(* IEC 61131-3 sources: 2026_Projet_YGO_ExcavatriceDragage/ARCHIVES/Code/PLC_TESTS, 2 files *)

(* ---- GVL_PLC_Tests_Const.st ---- *)
(* ═══════════════════════════════════════════════════════════════
   🧪 GVL_PLC_Tests_Const — Constantes de dimensionnement
   ───────────────────────────────────────────────────────────────
   🎯 Rôle : Définit les tailles limites des tables de tests
      pour l'orchestrateur et le moteur de tests.
   ═══════════════════════════════════════════════════════════════ *)

{attribute 'qualified_only'}
VAR_GLOBAL CONSTANT
    MaxTestCases     : INT := 8;    // par suite
    MaxSteps         : INT := 128;  // par suite, table PLATE ; WINCH-CORE-01 ajoute les étapes 65..111
    MaxChecks        : INT := 64;   // CheckTable par suite
    MaxChecksPerStep : INT := 10;
    MaxInvariants    : INT := 4;    // actifs en parallèle
    MaxProbeBool     : INT := 32;
    MaxProbeDint     : INT := 16;    // INT/WORD/étapes séquenceur → conversion au câblage (WORD_TO_DINT)
    MaxProbeReal     : INT := 16;    // analogiques + TIME → REAL ms
    MaxAnalogStims   : INT := 4;    // instances FB_TestStimulus par suite
    MaxSeqValues     : INT := 8;    // plus gros poste mémoire par stim
    TaskCycleMs      : INT := 10;   // MainTask — base des mesures en cycles
    MaxSuiteDurationMs : DINT := 180000; // 🛡️ garde-fou orchestrateur : 3 min maximum par suite
    MaxTestEvents    : INT := 32;   // journal circulaire des événements
    SuiteSafety      : INT := 1;    // index de suite (Cmd.RunSuite)
    SuiteTranslation : INT := 2;    // index de suite Translation M3 (Cmd.RunSuite)
    SuiteBucket      : INT := 3;    // index de suite Bucket (Cmd.RunSuite)
    SuiteEncoder     : INT := 4;    // index de suite Codeurs/Homing nominal (Cmd.RunSuite)
    SuiteModes       : INT := 5;    // index de suite Modes/Homme-mort, post-suppression IHM_MANU (Cmd.RunSuite)
    SuiteHeartbeat   : INT := 6;    // index de suite Heartbeat IHM↔PLC (Cmd.RunSuite)
    SuiteSupervision : INT := 8;    // index Supervision/Persistance config — 7 = Framework Validation
END_VAR

(* ---- FB_TestSequencer.st ---- *)
FUNCTION_BLOCK FB_TestSequencer
VAR_INPUT
    Start       : BOOL;              // Front : lance la suite
    Abort       : BOOL;              // Niveau : arrêt immédiat propre
    CaseId      : INT;               // 0=tous ; 1..MaxTestCases=cas ciblé
END_VAR
VAR_IN_OUT                           // 🔗 zéro copie
    StepTable      : ARRAY[1..GVL_PLC_Tests_Const.MaxSteps]      OF ST_TestStepConfig;
    CheckTable     : ARRAY[1..GVL_PLC_Tests_Const.MaxChecks]     OF ST_TestCheckConfig;
    CaseTable      : ARRAY[1..GVL_PLC_Tests_Const.MaxTestCases]  OF ST_TestCaseConfig;
    InvariantTable : ARRAY[1..GVL_PLC_Tests_Const.MaxInvariants] OF ST_TestInvariantConfig;
    ProbeBool      : ARRAY[1..GVL_PLC_Tests_Const.MaxProbeBool]  OF BOOL;
    ProbeDint      : ARRAY[1..GVL_PLC_Tests_Const.MaxProbeDint]  OF DINT;
    ProbeReal      : ARRAY[1..GVL_PLC_Tests_Const.MaxProbeReal]  OF REAL;
    Report         : ST_TestSuiteReport;
END_VAR
VAR_OUTPUT
    Busy                : BOOL;
    Done                : BOOL;
    AnyFailed           : BOOL;
    ConfigError         : BOOL;      // 🔒 Table invalide -> refus de lancer
    ConfigErrorStepId   : INT;
    ConfigErrorCheckIdx : INT;
    TerminalState       : E_TestTerminalState;
    ErrorCode           : INT;
    ErrorMessage        : STRING(160);
    CurrentStepId       : INT;
    ActiveStimulusId    : INT;       // ⚡ consommé par le domaine
    StepElapsed         : TIME;      // Pour l'IHM
END_VAR
VAR
    StartTrig           : R_TRIG;
    StepTimer           : TON;
    DwellTimer          : TON;
    Checks              : ARRAY[1..GVL_PLC_Tests_Const.MaxChecksPerStep] OF FB_TestCheck;
    InvChecks           : ARRAY[1..GVL_PLC_Tests_Const.MaxInvariants]    OF FB_TestCheck;
    InvArmed            : ARRAY[1..GVL_PLC_Tests_Const.MaxInvariants]    OF BOOL;

    // Variables de contrôle internes
    StepStarted         : BOOL;
    CurrentCaseId       : INT;
    Idx                 : INT;
    Jdx                 : INT;
    Kdx                 : INT;
    Valid               : BOOL;

    // 🔧 REX : locaux remontés depuis des blocs VAR imbriqués dans le corps
    AllChecksPassed     : BOOL;
    AnyCheckFailed      : BOOL;
    FailedCheckIdxLocal : INT;
    FailReasonLocal     : E_TestFailReason;
    ObsBoolLocal        : BOOL;
    ObsDintLocal        : DINT;
    ObsRealLocal        : REAL;
    NeverDuringPassed   : BOOL;
    SuiteAllPassed      : BOOL;
    FirstFailedCase     : INT;
    CaseIdx             : INT;
    CaseStartStep       : INT;
    CaseStep            : INT;
    CaseWalkCount       : INT;
    CaseOk              : BOOL;
    CaseExecuted        : BOOL;
    CaseFailedStep      : INT;
    CaseDuration        : TIME;
    CaseFailReason      : E_TestFailReason;

    // 🏷️ Construction de Report.FailureSummary (1 ligne lisible, tous les cas en échec)
    ReasonText          : STRING(20);
    EntryText           : STRING(80);
    FirstStepLocal      : INT;
    RequestedCaseId     : INT;
END_VAR
// === IMPLEMENTATION ===
StartTrig(CLK := Start);

// 1. Validation de la configuration sur front de Start
IF StartTrig.Q THEN
    ConfigError := FALSE;
    ConfigErrorStepId := 0;
    ConfigErrorCheckIdx := 0;
    TerminalState := E_TestTerminalState.TEST_TERMINAL_NONE;
    ErrorCode := 0;
    ErrorMessage := '';

    // 🛡️ Résolution interne CaseId → première étape, jamais d'étape exposée.
    RequestedCaseId := CaseId;
    IF CaseId < 0 OR CaseId > GVL_PLC_Tests_Const.MaxTestCases THEN
        ConfigError := TRUE;
        ConfigErrorStepId := CaseId;
        ErrorCode := 1001;
        ErrorMessage := 'CaseId hors limites';
        FirstStepLocal := 0;
    ELSIF CaseId = 0 THEN
        FirstStepLocal := CaseTable[1].FirstStep;
    ELSE
        FirstStepLocal := CaseTable[CaseId].FirstStep;
    END_IF;
    IF NOT ConfigError THEN
        IF FirstStepLocal < 1 OR FirstStepLocal > GVL_PLC_Tests_Const.MaxSteps THEN
            ConfigError := TRUE;
            ConfigErrorStepId := FirstStepLocal;
            ErrorCode := 1001;
            ErrorMessage := 'CaseTable.FirstStep hors limites';
        END_IF;
    END_IF;

    // Validation des étapes
    FOR Idx := 1 TO GVL_PLC_Tests_Const.MaxSteps DO
        IF StepTable[Idx].CaseId > 0 THEN
            // Vérification des NextOn
            IF StepTable[Idx].NextOnPass < 0 OR StepTable[Idx].NextOnPass > GVL_PLC_Tests_Const.MaxSteps THEN
                ConfigError := TRUE;
                ConfigErrorStepId := Idx;
            ELSIF StepTable[Idx].NextOnFail < 0 OR StepTable[Idx].NextOnFail > GVL_PLC_Tests_Const.MaxSteps THEN
                ConfigError := TRUE;
                ConfigErrorStepId := Idx;
            END_IF;

            // Vérification du Timeout
            IF StepTable[Idx].TimeoutPT <= T#0s THEN
                // Sauf si tous les checks de cette étape sont NEVER_DURING, mais restons stricts : TimeoutPT requis
                ConfigError := TRUE;
                ConfigErrorStepId := Idx;
            END_IF;

            // Vérification des Checks indexés par l'étape
            FOR Jdx := 1 TO GVL_PLC_Tests_Const.MaxChecksPerStep DO
                Kdx := StepTable[Idx].CheckIdx[Jdx];
                IF Kdx > 0 THEN
                    IF Kdx > GVL_PLC_Tests_Const.MaxChecks THEN
                        ConfigError := TRUE;
                        ConfigErrorStepId := Idx;
                        ConfigErrorCheckIdx := Kdx;
                    ELSE
                        // Validation de la sonde associée au check
                        CASE CheckTable[Kdx].Kind OF
                            E_TestCheckKind.BOOL_EQUAL, E_TestCheckKind.BOOL_RISING, E_TestCheckKind.BOOL_FALLING:
                                IF CheckTable[Kdx].ProbeIdx < 1 OR CheckTable[Kdx].ProbeIdx > GVL_PLC_Tests_Const.MaxProbeBool THEN
                                    ConfigError := TRUE;
                                    ConfigErrorStepId := Idx;
                                    ConfigErrorCheckIdx := Kdx;
                                END_IF;
                            E_TestCheckKind.DINT_EQUAL, E_TestCheckKind.DINT_NOT_EQUAL, E_TestCheckKind.DINT_IN_RANGE,
                            E_TestCheckKind.WORD_MASK_ALL, E_TestCheckKind.WORD_MASK_ANY, E_TestCheckKind.WORD_MASK_NONE:
                                IF CheckTable[Kdx].ProbeIdx < 1 OR CheckTable[Kdx].ProbeIdx > GVL_PLC_Tests_Const.MaxProbeDint THEN
                                    ConfigError := TRUE;
                                    ConfigErrorStepId := Idx;
                                    ConfigErrorCheckIdx := Kdx;
                                END_IF;
                            E_TestCheckKind.REAL_IN_RANGE:
                                IF CheckTable[Kdx].ProbeIdx < 1 OR CheckTable[Kdx].ProbeIdx > GVL_PLC_Tests_Const.MaxProbeReal THEN
                                    ConfigError := TRUE;
                                    ConfigErrorStepId := Idx;
                                    ConfigErrorCheckIdx := Kdx;
                                END_IF;
                        END_CASE;
                    END_IF;
                END_IF;
            END_FOR;
        END_IF;
    END_FOR;

    // 🛡️ ConfigError doit toujours produire Done + un état terminal.
    IF ConfigError THEN
        Busy := FALSE;
        Done := TRUE;
        AnyFailed := TRUE;
        ActiveStimulusId := 0;
        CurrentStepId := 0;
        StepElapsed := T#0s;
        TerminalState := E_TestTerminalState.TEST_TERMINAL_CONFIG_ERROR;
        Report.InProgress := FALSE;
        Report.RunCounter := Report.RunCounter + 1;
        Report.AllPassed := FALSE;
        Report.AnyFailed := TRUE;
        Report.Aborted := FALSE;
        Report.TerminalState := TerminalState;
        IF ErrorCode = 0 THEN
            ErrorCode := 1002;
            ErrorMessage := 'Table de test invalide';
        END_IF;
        Report.ErrorCode := ErrorCode;
        Report.ErrorMessage := ErrorMessage;
        Report.FailureSummary := CONCAT('CONFIG_ERROR step ', INT_TO_STRING(ConfigErrorStepId));
        RETURN;
    END_IF;
END_IF;

// 2. Abort (Niveau, priorité absolue)
IF Abort THEN
    IF Busy THEN
        Report.InProgress := FALSE;
        Report.Aborted := TRUE;
        Report.AnyFailed := TRUE;

        // Enregistrement de l'échec de l'étape courante
        IF CurrentStepId >= 1 AND CurrentStepId <= GVL_PLC_Tests_Const.MaxSteps THEN
            Report.Steps[CurrentStepId].Executed := TRUE;
            Report.Steps[CurrentStepId].Passed := FALSE;
            Report.Steps[CurrentStepId].FailReason := E_TestFailReason.FAIL_ABORTED;
            Report.Steps[CurrentStepId].Duration := StepElapsed;
        END_IF;

        // Échec du cas de test en cours
        IF CurrentCaseId >= 1 AND CurrentCaseId <= GVL_PLC_Tests_Const.MaxTestCases THEN
            Report.Cases[CurrentCaseId].Ok := FALSE;
            Report.Cases[CurrentCaseId].FailReason := E_TestFailReason.FAIL_ABORTED;
        END_IF;

        Busy := FALSE;
        Done := TRUE;
        AnyFailed := TRUE;
        TerminalState := E_TestTerminalState.TEST_TERMINAL_ABORTED;
        Report.TerminalState := TerminalState;
    END_IF;
    ActiveStimulusId := 0;
    StepStarted := FALSE;
    RETURN;
END_IF;

// 3. Démarrage de la suite
IF StartTrig.Q AND NOT ConfigError THEN
    Busy := TRUE;
    Done := FALSE;
    AnyFailed := FALSE;
    CurrentStepId := FirstStepLocal;
    StepStarted := FALSE;

    // RAZ Rapport
    Report.InProgress := TRUE;
    Report.AllPassed := FALSE;
    Report.AnyFailed := FALSE;
    Report.Aborted := FALSE;
    Report.TerminalState := E_TestTerminalState.TEST_TERMINAL_NONE;
    Report.ErrorCode := 0;
    Report.ErrorMessage := '';
    Report.FailedTestCase := 0;
    Report.CurrentStepId := FirstStepLocal;
    IF CurrentStepId >= 1 AND CurrentStepId <= GVL_PLC_Tests_Const.MaxSteps THEN
        Report.CurrentCaseId := StepTable[CurrentStepId].CaseId;
    ELSE
        Report.CurrentCaseId := 0;
    END_IF;
    Report.Duration := T#0s;
    Report.RunCounter := Report.RunCounter + 1;

    FOR Idx := 1 TO GVL_PLC_Tests_Const.MaxSteps DO
        Report.Steps[Idx].Executed := FALSE;
        Report.Steps[Idx].Passed := FALSE;
        Report.Steps[Idx].FailReason := E_TestFailReason.FAIL_NONE;
        Report.Steps[Idx].FailedCheckIdx := 0;
        Report.Steps[Idx].FailedInvariantId := 0;
        Report.Steps[Idx].Duration := T#0s;
    END_FOR;

    FOR Idx := 1 TO GVL_PLC_Tests_Const.MaxTestCases DO
        Report.Cases[Idx].Executed := FALSE;
        Report.Cases[Idx].Ok := FALSE;
        Report.Cases[Idx].FailedStepId := 0;
        Report.Cases[Idx].FailReason := E_TestFailReason.FAIL_NONE;
        Report.Cases[Idx].Duration := T#0s;
    END_FOR;

    // RAZ Invariants
    FOR Idx := 1 TO GVL_PLC_Tests_Const.MaxInvariants DO
        InvArmed[Idx] := FALSE;
    END_FOR;
END_IF;

// 4. Moteur d'exécution principal
IF Busy THEN
    // Incrément de la durée globale du run
    Report.Duration := Report.Duration + UDINT_TO_TIME(INT_TO_UDINT(GVL_PLC_Tests_Const.TaskCycleMs));

    // Vérification des bornes de l'étape courante (0 est valide et désigne la fin)
    IF CurrentStepId <> 0 AND (CurrentStepId < 1 OR CurrentStepId > GVL_PLC_Tests_Const.MaxSteps) THEN
        Busy := FALSE;
        Done := TRUE;
        AnyFailed := TRUE;
        ActiveStimulusId := 0;
        ConfigError := TRUE;
        ConfigErrorStepId := CurrentStepId;
        ErrorCode := 1003;
        ErrorMessage := 'Etape courante hors limites';
        TerminalState := E_TestTerminalState.TEST_TERMINAL_CONFIG_ERROR;
        Report.InProgress := FALSE;
        Report.AnyFailed := TRUE;
        Report.TerminalState := TerminalState;
        Report.ErrorCode := ErrorCode;
        Report.ErrorMessage := ErrorMessage;
        Report.FailureSummary := ErrorMessage;
        RETURN;
    END_IF;

    // 🔒 Fin automatique dès qu'un run ciblé tenterait d'entrer dans le cas suivant.
    IF CurrentStepId > 0 AND RequestedCaseId > 0 THEN
        IF StepTable[CurrentStepId].CaseId <> RequestedCaseId THEN
            CurrentStepId := 0;
            ActiveStimulusId := 0;
            StepStarted := FALSE;
        END_IF;
    END_IF;

    IF CurrentStepId > 0 THEN
    CurrentCaseId := StepTable[CurrentStepId].CaseId;
    ActiveStimulusId := StepTable[CurrentStepId].StimulusId;
    Report.CurrentStepId := CurrentStepId;
    Report.CurrentCaseId := CurrentCaseId;

    IF NOT StepStarted THEN
        StepStarted := TRUE;
        StepElapsed := T#0s;
        DwellTimer(IN := FALSE);
        StepTimer(IN := FALSE);

        // Gestion de l'armement/désarmement des invariants
        FOR Idx := 1 TO GVL_PLC_Tests_Const.MaxInvariants DO
            IF InvariantTable[Idx].ArmAtStepId = CurrentStepId THEN
                InvArmed[Idx] := TRUE;
            END_IF;
            IF InvariantTable[Idx].DisarmAtStepId = CurrentStepId THEN
                InvArmed[Idx] := FALSE;
            END_IF;
        END_FOR;
    END_IF;

    // Incrément de la durée de l'étape courante
    StepElapsed := StepElapsed + UDINT_TO_TIME(INT_TO_UDINT(GVL_PLC_Tests_Const.TaskCycleMs));

    // 4.1 Évaluation des invariants actifs
    FOR Idx := 1 TO GVL_PLC_Tests_Const.MaxInvariants DO
        IF InvArmed[Idx] THEN
            InvChecks[Idx](Config := InvariantTable[Idx].Check, Evaluate := TRUE, ProbeBool := ProbeBool, ProbeDint := ProbeDint, ProbeReal := ProbeReal);
            IF InvChecks[Idx].Failed THEN
                // Violation d'invariant -> Transition en échec immédiat
                Report.Steps[CurrentStepId].Executed := TRUE;
                Report.Steps[CurrentStepId].Passed := FALSE;
                Report.Steps[CurrentStepId].FailReason := E_TestFailReason.FAIL_INVARIANT;
                Report.Steps[CurrentStepId].FailedInvariantId := Idx;
                Report.Steps[CurrentStepId].Duration := StepElapsed;
                Report.Steps[CurrentStepId].ObservedBool := InvChecks[Idx].ObservedBool;
                Report.Steps[CurrentStepId].ObservedDint := InvChecks[Idx].ObservedDint;
                Report.Steps[CurrentStepId].ObservedReal := InvChecks[Idx].ObservedReal;

                // Désactivation de l'évaluation
                InvChecks[Idx](Config := InvariantTable[Idx].Check, Evaluate := FALSE, ProbeBool := ProbeBool, ProbeDint := ProbeDint, ProbeReal := ProbeReal);

                // Transition
                IF StepTable[CurrentStepId].FailAction = E_TestFailAction.FAIL_ABORT_SUITE THEN
                    Busy := FALSE;
                    Done := TRUE;
                    AnyFailed := TRUE;
                    ActiveStimulusId := 0;
                ELSE
                    CurrentStepId := StepTable[CurrentStepId].NextOnFail;
                    StepStarted := FALSE;
                END_IF;
                RETURN;
            END_IF;
        END_IF;
    END_FOR;

    // 4.2 Gestion de la temporisation de Dwell
    DwellTimer(IN := TRUE, PT := StepTable[CurrentStepId].DwellPT);
    IF NOT DwellTimer.Q THEN
        // En attente du Dwell, pas d'évaluation des checks d'étape
        FOR Jdx := 1 TO GVL_PLC_Tests_Const.MaxChecksPerStep DO
            Checks[Jdx](Evaluate := FALSE, ProbeBool := ProbeBool, ProbeDint := ProbeDint, ProbeReal := ProbeReal);
        END_FOR;
        RETURN;
    END_IF;

    // 4.3 Évaluation des checks d'étape
    AllChecksPassed     := TRUE;
    AnyCheckFailed      := FALSE;
    FailedCheckIdxLocal := 0;
    FailReasonLocal     := E_TestFailReason.FAIL_NONE;
    ObsBoolLocal        := FALSE;
    ObsDintLocal        := 0;
    ObsRealLocal        := 0.0;

    FOR Jdx := 1 TO GVL_PLC_Tests_Const.MaxChecksPerStep DO
        Kdx := StepTable[CurrentStepId].CheckIdx[Jdx];
        IF Kdx < 0 OR Kdx > GVL_PLC_Tests_Const.MaxChecks THEN
            ConfigError := TRUE;
            ConfigErrorStepId := CurrentStepId;
            ConfigErrorCheckIdx := Kdx;
            ErrorCode := 1006;
            ErrorMessage := 'CheckIdx runtime hors limites';
            Busy := FALSE;
            Done := TRUE;
            AnyFailed := TRUE;
            ActiveStimulusId := 0;
            TerminalState := E_TestTerminalState.TEST_TERMINAL_CONFIG_ERROR;
            RETURN;
        END_IF;
        IF Kdx > 0 THEN
            Checks[Jdx](Config := CheckTable[Kdx], Evaluate := TRUE, ProbeBool := ProbeBool, ProbeDint := ProbeDint, ProbeReal := ProbeReal);

            IF Checks[Jdx].Failed THEN
                AnyCheckFailed := TRUE;
                FailedCheckIdxLocal := Kdx;
                FailReasonLocal := Checks[Jdx].FailReason;
                ObsBoolLocal := Checks[Jdx].ObservedBool;
                ObsDintLocal := Checks[Jdx].ObservedDint;
                ObsRealLocal := Checks[Jdx].ObservedReal;
            ELSIF Checks[Jdx].Pending THEN
                AllChecksPassed := FALSE;
            END_IF;
        END_IF;
    END_FOR;

    // 4.4 Prise de verdict
    IF AnyCheckFailed THEN
        // Échec sur un check d'étape
        Report.Steps[CurrentStepId].Executed := TRUE;
        Report.Steps[CurrentStepId].Passed := FALSE;
        Report.Steps[CurrentStepId].FailReason := FailReasonLocal;
        Report.Steps[CurrentStepId].FailedCheckIdx := FailedCheckIdxLocal;
        Report.Steps[CurrentStepId].Duration := StepElapsed;
        Report.Steps[CurrentStepId].ObservedBool := ObsBoolLocal;
        Report.Steps[CurrentStepId].ObservedDint := ObsDintLocal;
        Report.Steps[CurrentStepId].ObservedReal := ObsRealLocal;

        // Reset checks
        FOR Jdx := 1 TO GVL_PLC_Tests_Const.MaxChecksPerStep DO
            Checks[Jdx](Evaluate := FALSE, ProbeBool := ProbeBool, ProbeDint := ProbeDint, ProbeReal := ProbeReal);
        END_FOR;

        IF StepTable[CurrentStepId].FailAction = E_TestFailAction.FAIL_ABORT_SUITE THEN
            Busy := FALSE;
            Done := TRUE;
            AnyFailed := TRUE;
            ActiveStimulusId := 0;
        ELSE
            CurrentStepId := StepTable[CurrentStepId].NextOnFail;
            StepStarted := FALSE;
        END_IF;
        RETURN;
    END_IF;

    StepTimer(IN := TRUE, PT := StepTable[CurrentStepId].TimeoutPT);

    IF AllChecksPassed THEN
        // Succès précoce (vérification MinPT)
        IF StepElapsed < StepTable[CurrentStepId].MinPT THEN
            // Réaction trop rapide = Échec
            Report.Steps[CurrentStepId].Executed := TRUE;
            Report.Steps[CurrentStepId].Passed := FALSE;
            Report.Steps[CurrentStepId].FailReason := E_TestFailReason.FAIL_WINDOW_EARLY;
            Report.Steps[CurrentStepId].Duration := StepElapsed;

            // Reset checks
            FOR Jdx := 1 TO GVL_PLC_Tests_Const.MaxChecksPerStep DO
                Checks[Jdx](Evaluate := FALSE, ProbeBool := ProbeBool, ProbeDint := ProbeDint, ProbeReal := ProbeReal);
            END_FOR;

            IF StepTable[CurrentStepId].FailAction = E_TestFailAction.FAIL_ABORT_SUITE THEN
                Busy := FALSE;
                Done := TRUE;
                AnyFailed := TRUE;
                ActiveStimulusId := 0;
            ELSE
                CurrentStepId := StepTable[CurrentStepId].NextOnFail;
                StepStarted := FALSE;
            END_IF;
        ELSE
            // Validation étape OK
            Report.Steps[CurrentStepId].Executed := TRUE;
            Report.Steps[CurrentStepId].Passed := TRUE;
            Report.Steps[CurrentStepId].Duration := StepElapsed;

            // Prendre snapshot du premier check s'il existe
            IF StepTable[CurrentStepId].CheckIdx[1] > 0 THEN
                Report.Steps[CurrentStepId].ObservedBool := Checks[1].ObservedBool;
                Report.Steps[CurrentStepId].ObservedDint := Checks[1].ObservedDint;
                Report.Steps[CurrentStepId].ObservedReal := Checks[1].ObservedReal;
            END_IF;

            // Reset checks
            FOR Jdx := 1 TO GVL_PLC_Tests_Const.MaxChecksPerStep DO
                Checks[Jdx](Evaluate := FALSE, ProbeBool := ProbeBool, ProbeDint := ProbeDint, ProbeReal := ProbeReal);
            END_FOR;

            CurrentStepId := StepTable[CurrentStepId].NextOnPass;
            StepStarted := FALSE;
        END_IF;
        RETURN;
    END_IF;

    // Gestion du timeout d'étape
    IF StepTimer.Q THEN
        // Si timeout expiré, vérifions si des checks NEVER_DURING sont en attente
        NeverDuringPassed := TRUE;
        FOR Jdx := 1 TO GVL_PLC_Tests_Const.MaxChecksPerStep DO
            Kdx := StepTable[CurrentStepId].CheckIdx[Jdx];
            IF Kdx < 0 OR Kdx > GVL_PLC_Tests_Const.MaxChecks THEN
                ConfigError := TRUE;
                ConfigErrorStepId := CurrentStepId;
                ConfigErrorCheckIdx := Kdx;
                ErrorCode := 1006;
                ErrorMessage := 'CheckIdx timeout hors limites';
                Busy := FALSE;
                Done := TRUE;
                AnyFailed := TRUE;
                ActiveStimulusId := 0;
                TerminalState := E_TestTerminalState.TEST_TERMINAL_CONFIG_ERROR;
                RETURN;
            END_IF;
            IF Kdx > 0 THEN
                IF CheckTable[Kdx].Mode = E_TestCheckMode.CHECK_NEVER_DURING THEN
                    // Jamais violé pendant toute la fenêtre
                    Checks[Jdx](Evaluate := FALSE, ProbeBool := ProbeBool, ProbeDint := ProbeDint, ProbeReal := ProbeReal);
                ELSE
                    // Les autres modes auraient dû passer avant le timeout
                    NeverDuringPassed := FALSE;
                END_IF;
            END_IF;
        END_FOR;

        IF NeverDuringPassed THEN
            // Succès par non-violation
            Report.Steps[CurrentStepId].Executed := TRUE;
            Report.Steps[CurrentStepId].Passed := TRUE;
            Report.Steps[CurrentStepId].Duration := StepElapsed;

            CurrentStepId := StepTable[CurrentStepId].NextOnPass;
            StepStarted := FALSE;
        ELSE
            // Timeout classique de l'étape
            Report.Steps[CurrentStepId].Executed := TRUE;
            Report.Steps[CurrentStepId].Passed := FALSE;
            Report.Steps[CurrentStepId].FailReason := E_TestFailReason.FAIL_TIMEOUT;
            Report.Steps[CurrentStepId].Duration := StepElapsed;

            IF StepTable[CurrentStepId].FailAction = E_TestFailAction.FAIL_ABORT_SUITE THEN
                Busy := FALSE;
                Done := TRUE;
                AnyFailed := TRUE;
                ActiveStimulusId := 0;
            ELSE
                CurrentStepId := StepTable[CurrentStepId].NextOnFail;
                StepStarted := FALSE;
            END_IF;
        END_IF;

        // Reset checks
        FOR Jdx := 1 TO GVL_PLC_Tests_Const.MaxChecksPerStep DO
            Checks[Jdx](Evaluate := FALSE, ProbeBool := ProbeBool, ProbeDint := ProbeDint, ProbeReal := ProbeReal);
        END_FOR;
    END_IF;
    END_IF;
END_IF;

// 5. Agrégation des résultats en fin de suite (CurrentStepId = 0)
IF Busy AND CurrentStepId = 0 THEN
    Busy := FALSE;
    Done := TRUE;
    ActiveStimulusId := 0;
    Report.InProgress := FALSE;

    // Agrégation des cas de test
    SuiteAllPassed  := TRUE;
    FirstFailedCase := 0;

    FOR CaseIdx := 1 TO GVL_PLC_Tests_Const.MaxTestCases DO
        CaseStartStep := CaseTable[CaseIdx].FirstStep;
        IF CaseStartStep > 0 THEN
            CaseOk := TRUE;
            CaseExecuted := FALSE;
            CaseFailedStep := 0;
            CaseDuration := T#0s;
            CaseFailReason := E_TestFailReason.FAIL_NONE;

            // 🔒 Parcours borné et index validé AVANT déréférencement.
            // CODESYS peut évaluer StepTable[CaseStep] même si CaseStep=0
            // dans une condition composée : ancienne version = Access Violation CPU.
            CaseStep := CaseStartStep;
            FOR CaseWalkCount := 1 TO GVL_PLC_Tests_Const.MaxSteps DO
                IF CaseStep = 0 THEN
                    EXIT;
                END_IF;
                IF CaseStep < 1 OR CaseStep > GVL_PLC_Tests_Const.MaxSteps THEN
                    ConfigError := TRUE;
                    ConfigErrorStepId := CaseStep;
                    ErrorCode := 1004;
                    ErrorMessage := 'Agregation : etape hors limites';
                    CaseOk := FALSE;
                    EXIT;
                END_IF;
                IF StepTable[CaseStep].CaseId <> CaseIdx THEN
                    EXIT;
                END_IF;

                IF Report.Steps[CaseStep].Executed THEN
                    CaseExecuted := TRUE;
                    CaseDuration := CaseDuration + Report.Steps[CaseStep].Duration;
                    IF NOT Report.Steps[CaseStep].Passed THEN
                        CaseOk := FALSE;
                        CaseFailedStep := CaseStep;
                        CaseFailReason := Report.Steps[CaseStep].FailReason;
                        CaseStep := StepTable[CaseStep].NextOnFail;
                    ELSE
                        CaseStep := StepTable[CaseStep].NextOnPass;
                    END_IF;
                ELSE
                    CaseStep := StepTable[CaseStep].NextOnPass;
                END_IF;
            END_FOR;
            IF CaseStep <> 0 AND CaseWalkCount > GVL_PLC_Tests_Const.MaxSteps THEN
                ConfigError := TRUE;
                ConfigErrorStepId := CaseStep;
                ErrorCode := 1005;
                ErrorMessage := 'Agregation : cycle de transitions';
                CaseOk := FALSE;
            END_IF;

            Report.Cases[CaseIdx].Name := CaseTable[CaseIdx].Name; // 🏷️ Lisible directement en Watch, sans chercher l'index
            Report.Cases[CaseIdx].Executed := CaseExecuted;
            Report.Cases[CaseIdx].Ok := CaseExecuted AND CaseOk;
            Report.Cases[CaseIdx].FailedStepId := CaseFailedStep;
            Report.Cases[CaseIdx].FailReason := CaseFailReason;
            Report.Cases[CaseIdx].Duration := CaseDuration;

            IF CaseExecuted AND NOT CaseOk THEN
                SuiteAllPassed := FALSE;
                IF FirstFailedCase = 0 THEN
                    FirstFailedCase := CaseIdx;
                END_IF;
            END_IF;
        END_IF;
    END_FOR;

    Report.AllPassed := SuiteAllPassed;
    Report.AnyFailed := NOT SuiteAllPassed;
    Report.FailedTestCase := FirstFailedCase;
    AnyFailed := NOT SuiteAllPassed;
    IF SuiteAllPassed THEN
        TerminalState := E_TestTerminalState.TEST_TERMINAL_DONE;
    ELSE
        TerminalState := E_TestTerminalState.TEST_TERMINAL_FAILED;
    END_IF;
    Report.TerminalState := TerminalState;
    Report.ErrorCode := ErrorCode;
    Report.ErrorMessage := ErrorMessage;

    // 🏷️ Résumé texte de TOUS les cas en échec (pas juste le premier) — évite de
    // parcourir Cases[] un par un en Watch (demande utilisateur 2026-07-16)
    Report.FailureSummary := '';
    FOR CaseIdx := 1 TO GVL_PLC_Tests_Const.MaxTestCases DO
        IF Report.Cases[CaseIdx].Executed AND NOT Report.Cases[CaseIdx].Ok THEN
            CASE Report.Cases[CaseIdx].FailReason OF
                E_TestFailReason.FAIL_TIMEOUT:      ReasonText := 'FAIL_TIMEOUT';
                E_TestFailReason.FAIL_CHECK:        ReasonText := 'FAIL_CHECK';
                E_TestFailReason.FAIL_INVARIANT:    ReasonText := 'FAIL_INVARIANT';
                E_TestFailReason.FAIL_WINDOW_EARLY: ReasonText := 'FAIL_WINDOW_EARLY';
                E_TestFailReason.FAIL_ABORTED:      ReasonText := 'FAIL_ABORTED';
            ELSE
                ReasonText := 'FAIL_NONE';
            END_CASE;

            EntryText := CONCAT(Report.Cases[CaseIdx].Name, ' (step ');
            EntryText := CONCAT(EntryText, INT_TO_STRING(Report.Cases[CaseIdx].FailedStepId));
            EntryText := CONCAT(EntryText, '): ');
            EntryText := CONCAT(EntryText, ReasonText);

            IF Report.FailureSummary = '' THEN
                Report.FailureSummary := EntryText;
            ELSE
                Report.FailureSummary := CONCAT(Report.FailureSummary, ' | ');
                Report.FailureSummary := CONCAT(Report.FailureSummary, EntryText);
            END_IF;
        END_IF;
    END_FOR;
END_IF;
